// TIA Portal V14 SP1 export
// export: Created 2000-01-01T00:00:00.0000000Z, ExportSetting WithDefaults, WithReadOnly
TYPE "MCP_RC_UDT"
   STRUCT
      Run : Bool;   // Run command
      Speed : Int;
   END_STRUCT;
END_TYPE
